      FC_W[1,14] := 0.00180894;
      FC_W[1,15] := -1.01147878;
      FC_W[1,16] := 0.31076741;
      FC_W[1,17] := -0.42154586;
      FC_W[1,18] := -0.05431300;
      FC_W[1,19] := 0.68237108;
      FC_W[1,20] := -2.56503296;
      FC_W[1,21] := 0.50673449;
      FC_W[1,22] := 0.31768897;
      FC_W[1,23] := -0.43834999;
      FC_W[1,24] := 1.20007265;
      FC_W[1,25] := 0.30830422;
      FC_W[1,26] := 0.13145778;
      FC_W[1,27] := 0.41129708;
      FC_W[1,28] := -0.09861557;
      FC_W[1,29] := -0.05401544;
      FC_W[1,30] := -0.38849521;
      FC_W[1,31] := -1.97921050;
      FC_W[2,0] := -0.79939067;
      FC_W[2,1] := 0.10302242;
      FC_W[2,2] := 0.09020624;
      FC_W[2,3] := -0.46045631;
      FC_W[2,4] := 0.32426205;
      FC_W[2,5] := 0.07683180;
      FC_W[2,6] := 0.54684573;
      FC_W[2,7] := 1.87505293;
      FC_W[2,8] := -0.48562393;
      FC_W[2,9] := 0.99263871;
      FC_W[2,10] := -0.65771282;
      FC_W[2,11] := 0.72155434;
      FC_W[2,12] := -0.66074061;
      FC_W[2,13] := 0.11306432;
      FC_W[2,14] := -0.38545227;
      FC_W[2,15] := 0.16300759;
      FC_W[2,16] := -0.02957736;
      FC_W[2,17] := -0.82533288;
      FC_W[2,18] := 0.33957723;
      FC_W[2,19] := -0.78074455;
      FC_W[2,20] := 0.55624270;
      FC_W[2,21] := -0.52731699;
      FC_W[2,22] := -1.25810063;
      FC_W[2,23] := -0.21556486;
      FC_W[2,24] := -0.03355473;
      FC_W[2,25] := 0.02170837;
      FC_W[2,26] := -0.12119742;
      FC_W[2,27] := -0.88717794;
      FC_W[2,28] := -0.91240627;
      FC_W[2,29] := 0.36170098;
      FC_W[2,30] := 0.16164558;
      FC_W[2,31] := 0.99094546;
      FC_W[3,0] := 0.19523349;
      FC_W[3,1] := 0.31197101;
      FC_W[3,2] := -0.48878455;
      FC_W[3,3] := 0.14373684;
      FC_W[3,4] := 0.24886017;
      FC_W[3,5] := -0.42134193;
      FC_W[3,6] := -0.14882350;
      FC_W[3,7] := 0.79451615;
      FC_W[3,8] := -0.46309730;
      FC_W[3,9] := 0.40033284;
      FC_W[3,10] := -0.68702614;
      FC_W[3,11] := -0.29239723;
      FC_W[3,12] := 0.98389262;
      FC_W[3,13] := 0.30846006;
      FC_W[3,14] := -0.12699004;
      FC_W[3,15] := 1.25244427;
      FC_W[3,16] := 0.17832240;
      FC_W[3,17] := -0.43285766;
      FC_W[3,18] := 0.26159754;
      FC_W[3,19] := 0.15949164;
      FC_W[3,20] := 1.06185210;
      FC_W[3,21] := 0.14212017;
      FC_W[3,22] := 0.00880439;
      FC_W[3,23] := -0.36065376;
      FC_W[3,24] := -0.39496204;
      FC_W[3,25] := -0.00392890;
      FC_W[3,26] := -0.77206844;
      FC_W[3,27] := -0.12771720;
      FC_W[3,28] := 0.72197872;
      FC_W[3,29] := 0.24183723;
      FC_W[3,30] := -0.38839531;
      FC_W[3,31] := 0.04649191;
      FC_W[4,0] := -0.42976218;
      FC_W[4,1] := 0.71019524;
      FC_W[4,2] := 0.02715457;
      FC_W[4,3] := 0.20727751;
      FC_W[4,4] := 0.12750632;
      FC_W[4,5] := 0.10362761;
      FC_W[4,6] := 0.56926334;
      FC_W[4,7] := 0.33267853;
      FC_W[4,8] := 0.22530533;
      FC_W[4,9] := -0.76057816;
      FC_W[4,10] := 0.06259055;
      FC_W[4,11] := 0.65855861;
      FC_W[4,12] := 0.43817779;
      FC_W[4,13] := -1.45052433;
      FC_W[4,14] := -0.69694483;
      FC_W[4,15] := 0.39829472;
      FC_W[4,16] := 0.00987289;
      FC_W[4,17] := 0.68149745;
      FC_W[4,18] := -0.59120047;
      FC_W[4,19] := 0.11526035;
      FC_W[4,20] := -0.45347911;
      FC_W[4,21] := 0.55277812;
      FC_W[4,22] := -0.36495659;
      FC_W[4,23] := -0.65428317;
      FC_W[4,24] := -2.59415770;
      FC_W[4,25] := 0.01274597;
      FC_W[4,26] := -0.42365780;
      FC_W[4,27] := 0.38587591;
      FC_W[4,28] := 0.33021146;
      FC_W[4,29] := 0.45073530;
      FC_W[4,30] := -0.22007711;
      FC_W[4,31] := 0.46025163;
      FC_W[5,0] := 0.08847263;
      FC_W[5,1] := 2.92971921;
      FC_W[5,2] := 0.40630540;
      FC_W[5,3] := -0.18477380;
      FC_W[5,4] := -0.35985741;
      FC_W[5,5] := 0.16343132;
      FC_W[5,6] := -1.01463449;
      FC_W[5,7] := -0.19884980;
      FC_W[5,8] := 0.19642729;
      FC_W[5,9] := 0.07467357;
      FC_W[5,10] := -0.20739354;
      FC_W[5,11] := -0.32682586;
      FC_W[5,12] := -0.24732944;
      FC_W[5,13] := -0.28553879;
      FC_W[5,14] := 0.02577983;
      FC_W[5,15] := -0.35895699;
      FC_W[5,16] := 0.13909405;
      FC_W[5,17] := -0.85842067;
      FC_W[5,18] := 0.29272711;
      FC_W[5,19] := 0.14367910;
      FC_W[5,20] := -0.33554327;
      FC_W[5,21] := -0.10857771;
      FC_W[5,22] := 0.06511363;
      FC_W[5,23] := 1.53560221;
      FC_W[5,24] := 0.36751866;
      FC_W[5,25] := 0.14096503;
      FC_W[5,26] := 0.68856186;
      FC_W[5,27] := -0.00372456;
      FC_W[5,28] := 0.07267709;
      FC_W[5,29] := 0.29737416;
      FC_W[5,30] := 0.05855417;
      FC_W[5,31] := 0.18817970;
      FC_W[6,0] := 0.22961207;
      FC_W[6,1] := 1.10309398;
      FC_W[6,2] := 1.14253712;
      FC_W[6,3] := -0.24431218;
      FC_W[6,4] := 0.24880899;
      FC_W[6,5] := 0.10031620;
      FC_W[6,6] := -1.37900984;
      FC_W[6,7] := -0.46621767;
      FC_W[6,8] := 0.23081133;
      FC_W[6,9] := -0.62265766;
      FC_W[6,10] := -0.19415495;
      FC_W[6,11] := 0.24065939;
      FC_W[6,12] := -0.37324443;
      FC_W[6,13] := 0.04941022;
      FC_W[6,14] := -0.58380717;
      FC_W[6,15] := 0.29722652;
      FC_W[6,16] := 0.45706749;
      FC_W[6,17] := 0.79749161;
      FC_W[6,18] := 0.24645862;
      FC_W[6,19] := -0.69690132;
      FC_W[6,20] := 0.25755104;
      FC_W[6,21] := -1.28122711;
      FC_W[6,22] := -0.90884095;
      FC_W[6,23] := -1.13884628;
      FC_W[6,24] := 0.61092412;
      FC_W[6,25] := 0.10356417;
      FC_W[6,26] := -0.16909865;
      FC_W[6,27] := -0.64685744;
      FC_W[6,28] := 0.09836304;
      FC_W[6,29] := 0.29990685;
      FC_W[6,30] := -0.26579708;
      FC_W[6,31] := -0.09385087;
      FC_W[7,0] := 0.11735278;
      FC_W[7,1] := 0.69732809;
      FC_W[7,2] := -0.28756016;
      FC_W[7,3] := -0.12583709;
      FC_W[7,4] := -0.44791237;
      FC_W[7,5] := 0.04257831;
      FC_W[7,6] := 0.01414247;
      FC_W[7,7] := 0.31274548;
      FC_W[7,8] := -0.42705598;
      FC_W[7,9] := 0.25311053;
      FC_W[7,10] := -0.02971629;
      FC_W[7,11] := 0.08217675;
      FC_W[7,12] := 1.13895476;
      FC_W[7,13] := 0.28638309;
      FC_W[7,14] := 0.30324531;
      FC_W[7,15] := 1.06351733;
      FC_W[7,16] := -0.09911025;
      FC_W[7,17] := -0.12825158;
      FC_W[7,18] := -0.21037468;
      FC_W[7,19] := -0.15125044;
      FC_W[7,20] := 1.04692757;
      FC_W[7,21] := -0.19273317;
      FC_W[7,22] := -0.01566108;
      FC_W[7,23] := -0.82813007;
      FC_W[7,24] := -0.17457560;
      FC_W[7,25] := -0.23310129;
      FC_W[7,26] := -0.67900503;
      FC_W[7,27] := -0.00216983;
      FC_W[7,28] := -0.33897799;
      FC_W[7,29] := 0.23453975;
      FC_W[7,30] := 0.43223280;
      FC_W[7,31] := 0.38816142;
      FC_W[8,0] := 1.24795640;
      FC_W[8,1] := 0.16966595;
      FC_W[8,2] := -0.59130764;
      FC_W[8,3] := -1.17259443;
      FC_W[8,4] := 0.58706713;
      FC_W[8,5] := -0.50881100;
      FC_W[8,6] := -0.93378001;
      FC_W[8,7] := 1.83182466;
      FC_W[8,8] := 0.69100636;
      FC_W[8,9] := -0.18218489;
      FC_W[8,10] := 0.03764156;
      FC_W[8,11] := -0.73455888;
      FC_W[8,12] := -0.53293765;
      FC_W[8,13] := 0.35738659;
      FC_W[8,14] := 0.34333083;
      FC_W[8,15] := 0.42288589;
      FC_W[8,16] := 0.47547165;
      FC_W[8,17] := 0.63862199;
      FC_W[8,18] := 0.62496924;
      FC_W[8,19] := 0.38435844;
      FC_W[8,20] := 1.82490015;
      FC_W[8,21] := 0.90129334;
      FC_W[8,22] := -0.10840212;
      FC_W[8,23] := 0.10254918;
      FC_W[8,24] := -0.91856247;
      FC_W[8,25] := 0.00505273;
      FC_W[8,26] := -0.97525537;
      FC_W[8,27] := 1.19635546;
      FC_W[8,28] := 0.29022071;
      FC_W[8,29] := 0.81490791;
      FC_W[8,30] := -0.35306564;
      FC_W[8,31] := -0.03846764;
      FC_W[9,0] := 0.53101271;
      FC_W[9,1] := 0.67765594;
      FC_W[9,2] := -0.31747413;
      FC_W[9,3] := -0.61590499;
      FC_W[9,4] := -0.35415921;
      FC_W[9,5] := 0.04045775;
      FC_W[9,6] := -0.25351635;
      FC_W[9,7] := 0.61500031;
      FC_W[9,8] := -0.00759591;
      FC_W[9,9] := 0.01995997;
      FC_W[9,10] := 0.31222284;
      FC_W[9,11] := -0.03113513;
      FC_W[9,12] := 0.55826259;
      FC_W[9,13] := 0.29481170;
      FC_W[9,14] := 0.50861734;
      FC_W[9,15] := 0.74235141;
      FC_W[9,16] := 0.04826086;
      FC_W[9,17] := 0.32700640;
      FC_W[9,18] := -0.14947560;
      FC_W[9,19] := -0.14729200;
      FC_W[9,20] := 1.31701505;
      FC_W[9,21] := 0.06887171;
      FC_W[9,22] := -0.09508032;
      FC_W[9,23] := -0.69279194;
      FC_W[9,24] := -0.32143742;
      FC_W[9,25] := -0.23362400;
      FC_W[9,26] := -0.77252012;
      FC_W[9,27] := 0.48929808;
      FC_W[9,28] := -0.59472609;
      FC_W[9,29] := 0.44059590;
      FC_W[9,30] := 0.51598865;
      FC_W[9,31] := 0.40399224;
      FC_W[10,0] := -0.05485313;
      FC_W[10,1] := 0.79143423;
      FC_W[10,2] := -0.47971761;
      FC_W[10,3] := -0.42792881;
      FC_W[10,4] := 0.76965564;
      FC_W[10,5] := 0.38477486;
      FC_W[10,6] := 0.42768925;
      FC_W[10,7] := 0.28604057;
      FC_W[10,8] := -1.25346828;
      FC_W[10,9] := 0.49736726;
      FC_W[10,10] := 0.69473928;
      FC_W[10,11] := 0.79891783;
      FC_W[10,12] := 0.62251019;
      FC_W[10,13] := 0.17432037;
      FC_W[10,14] := 1.53301835;
      FC_W[10,15] := 0.93965453;
      FC_W[10,16] := -0.46999088;
      FC_W[10,17] := 0.77361441;
      FC_W[10,18] := 0.22307561;
      FC_W[10,19] := -1.36293745;
      FC_W[10,20] := 0.20648916;
      FC_W[10,21] := 0.06673018;
      FC_W[10,22] := 0.22559744;
      FC_W[10,23] := 0.43268546;
      FC_W[10,24] := -0.21780904;
      FC_W[10,25] := -0.78115875;
      FC_W[10,26] := -0.24076101;
      FC_W[10,27] := 0.62123424;
      FC_W[10,28] := 0.29939529;
      FC_W[10,29] := 0.09014255;
      FC_W[10,30] := 0.25302246;
      FC_W[10,31] := -0.03954656;
      FC_W[11,0] := -0.24293564;
      FC_W[11,1] := -0.04531259;
      FC_W[11,2] := 0.00998670;
      FC_W[11,3] := 0.19956830;
      FC_W[11,4] := -0.20174095;
      FC_W[11,5] := -0.11596463;
      FC_W[11,6] := -0.22455990;
      FC_W[11,7] := -0.11557520;
      FC_W[11,8] := 0.41246292;
      FC_W[11,9] := 0.08150622;
      FC_W[11,10] := -1.95139670;
      FC_W[11,11] := -0.45480672;
      FC_W[11,12] := -0.08829422;
      FC_W[11,13] := 0.05833782;
      FC_W[11,14] := 0.26944444;
      FC_W[11,15] := 0.21539681;
      FC_W[11,16] := 2.23111510;
      FC_W[11,17] := 0.66294128;
      FC_W[11,18] := -0.05759437;
      FC_W[11,19] := -0.41524842;
      FC_W[11,20] := -0.13926855;
      FC_W[11,21] := 0.04841401;
      FC_W[11,22] := -0.05950727;
      FC_W[11,23] := 0.11197530;
      FC_W[11,24] := -0.04123791;
      FC_W[11,25] := -0.26082167;
      FC_W[11,26] := -0.45694438;
      FC_W[11,27] := 0.20621511;
      FC_W[11,28] := -0.53152508;
      FC_W[11,29] := 0.38166457;
      FC_W[11,30] := 0.31593123;
      FC_W[11,31] := 0.02903810;
      FC_W[12,0] := -0.11749745;
      FC_W[12,1] := -0.23415545;
      FC_W[12,2] := -0.34946913;
      FC_W[12,3] := 0.53356487;
      FC_W[12,4] := 0.18837753;
      FC_W[12,5] := -0.70393479;
      FC_W[12,6] := -0.50469047;
      FC_W[12,7] := -0.43645567;
      FC_W[12,8] := 0.66334420;
      FC_W[12,9] := -0.32834104;
      FC_W[12,10] := -1.24227428;
      FC_W[12,11] := -0.34643209;
      FC_W[12,12] := -0.28256458;
      FC_W[12,13] := -0.03548216;
      FC_W[12,14] := -0.02313955;
      FC_W[12,15] := 1.09937835;
      FC_W[12,16] := 1.40113294;
      FC_W[12,17] := 0.21808513;
      FC_W[12,18] := 0.18139383;
      FC_W[12,19] := -0.08548864;
      FC_W[12,20] := -0.56923884;
      FC_W[12,21] := 0.65053141;
      FC_W[12,22] := -0.65991580;
      FC_W[12,23] := 0.23657089;
      FC_W[12,24] := 0.02915133;
      FC_W[12,25] := -0.37136909;
      FC_W[12,26] := -0.20713671;
      FC_W[12,27] := 0.04201923;
      FC_W[12,28] := -0.21818402;
      FC_W[12,29] := 0.43879950;
      FC_W[12,30] := 0.66941983;
      FC_W[12,31] := 0.77976692;
      FC_W[13,0] := 0.05367998;
      FC_W[13,1] := 1.02593648;
      FC_W[13,2] := -1.72975278;
      FC_W[13,3] := 0.80966431;
      FC_W[13,4] := 0.03437574;
      FC_W[13,5] := -1.25336730;
      FC_W[13,6] := -0.54343611;
      FC_W[13,7] := -0.76846027;
      FC_W[13,8] := -0.07641880;
      FC_W[13,9] := -0.21239853;
      FC_W[13,10] := -1.32163453;
      FC_W[13,11] := 0.67327833;
      FC_W[13,12] := -1.27367902;
      FC_W[13,13] := -0.86751330;
      FC_W[13,14] := 0.55482459;
      FC_W[13,15] := -1.92334485;
      FC_W[13,16] := 0.08597323;
      FC_W[13,17] := -0.23974323;
      FC_W[13,18] := 0.09139446;
      FC_W[13,19] := 0.03227244;
      FC_W[13,20] := -0.22558706;
      FC_W[13,21] := -0.00554077;
      FC_W[13,22] := -0.24220449;
      FC_W[13,23] := -0.93250173;
      FC_W[13,24] := 1.33914196;
      FC_W[13,25] := -0.14073664;
      FC_W[13,26] := 1.38821757;
      FC_W[13,27] := -0.63530439;
      FC_W[13,28] := 0.86958200;
      FC_W[13,29] := -1.50805593;
      FC_W[13,30] := -0.21380891;
      FC_W[13,31] := 0.41014621;
      FC_W[14,0] := -0.63119894;
      FC_W[14,1] := -0.10577224;
      FC_W[14,2] := -0.08785659;
      FC_W[14,3] := -0.51354879;
      FC_W[14,4] := 0.30728057;
      FC_W[14,5] := -0.94762784;
      FC_W[14,6] := -0.00680102;
      FC_W[14,7] := 0.46720606;
      FC_W[14,8] := 2.24362016;
      FC_W[14,9] := -1.06858647;
      FC_W[14,10] := -1.56347978;
      FC_W[14,11] := -1.45889282;
      FC_W[14,12] := 0.46342093;
      FC_W[14,13] := 0.01371147;
      FC_W[14,14] := -0.43850195;
      FC_W[14,15] := -0.26042199;
      FC_W[14,16] := -2.62758970;
      FC_W[14,17] := -0.29780927;
      FC_W[14,18] := -1.96324050;
      FC_W[14,19] := -4.90748167;
      FC_W[14,20] := -0.20483738;
      FC_W[14,21] := -0.03886629;
      FC_W[14,22] := 1.46648896;
      FC_W[14,23] := 0.15051331;
      FC_W[14,24] := -0.04148193;
      FC_W[14,25] := -1.55939674;
      FC_W[14,26] := -0.01877716;
      FC_W[14,27] := -0.32644957;
      FC_W[14,28] := -0.03895755;
      FC_W[14,29] := -0.03125083;
      FC_W[14,30] := 0.01780568;
      FC_W[14,31] := -0.54571784;
      FC_W[15,0] := -0.89153206;
      FC_W[15,1] := 0.20046420;
      FC_W[15,2] := -0.15894163;
      FC_W[15,3] := -0.62003499;
      FC_W[15,4] := 0.67500734;
      FC_W[15,5] := -0.81095988;
      FC_W[15,6] := -0.43512601;
      FC_W[15,7] := 0.08051200;
      FC_W[15,8] := 0.22382137;
      FC_W[15,9] := 0.21324296;
      FC_W[15,10] := -1.19856393;
      FC_W[15,11] := -0.23485571;
      FC_W[15,12] := 0.08108855;
      FC_W[15,13] := -0.00869130;
      FC_W[15,14] := 0.20973921;
      FC_W[15,15] := -0.42064503;
      FC_W[15,16] := 0.83993143;
      FC_W[15,17] := 0.39107731;
      FC_W[15,18] := 0.05626461;
      FC_W[15,19] := 0.43600541;
      FC_W[15,20] := -0.40640157;
      FC_W[15,21] := -0.41479343;
      FC_W[15,22] := 1.18510294;
      FC_W[15,23] := 0.01747333;
      FC_W[15,24] := 0.27544057;
      FC_W[15,25] := 1.41735625;
      FC_W[15,26] := -1.28652883;
      FC_W[15,27] := -0.30560207;
      FC_W[15,28] := 0.28828090;
      FC_W[15,29] := 0.34294400;
      FC_W[15,30] := 1.56105816;
      FC_W[15,31] := 0.66715974;
      FC_W[16,0] := 0.18511236;
      FC_W[16,1] := 0.11142320;
      FC_W[16,2] := 0.25088802;
      FC_W[16,3] := 0.24562232;
      FC_W[16,4] := 0.23386742;
      FC_W[16,5] := 1.43394780;
      FC_W[16,6] := 1.17761219;
      FC_W[16,7] := -0.49213803;
      FC_W[16,8] := 1.12759876;
      FC_W[16,9] := 1.29781663;
      FC_W[16,10] := 0.37763405;
      FC_W[16,11] := -0.60559410;
      FC_W[16,12] := -0.58088464;
      FC_W[16,13] := -0.03103711;
      FC_W[16,14] := -0.37153244;
      FC_W[16,15] := 0.14177552;
      FC_W[16,16] := 0.08989498;
      FC_W[16,17] := -1.21121275;
      FC_W[16,18] := -1.52446818;
      FC_W[16,19] := -0.15327719;
      FC_W[16,20] := 1.36897111;
      FC_W[16,21] := -0.97303110;
      FC_W[16,22] := -1.61964941;
      FC_W[16,23] := -0.45303893;
      FC_W[16,24] := 0.07086476;
      FC_W[16,25] := -0.20691338;
      FC_W[16,26] := 0.56280392;
      FC_W[16,27] := 1.59726894;
      FC_W[16,28] := 3.60174441;
      FC_W[16,29] := -0.53792644;
      FC_W[16,30] := 2.29794812;
      FC_W[16,31] := -1.52492857;
      FC_W[17,0] := -1.34601951;
      FC_W[17,1] := -0.13013357;
      FC_W[17,2] := -0.39320931;
      FC_W[17,3] := -1.76083004;
      FC_W[17,4] := -0.25579280;
      FC_W[17,5] := -0.24240695;
      FC_W[17,6] := 0.40721077;
      FC_W[17,7] := -0.23947778;
      FC_W[17,8] := 0.50300777;
      FC_W[17,9] := -0.12915973;
      FC_W[17,10] := 3.87150478;
      FC_W[17,11] := 1.48434913;
      FC_W[17,12] := -0.27643603;
      FC_W[17,13] := 0.04503229;
      FC_W[17,14] := -0.24153562;
      FC_W[17,15] := -0.34765482;
      FC_W[17,16] := 2.79668903;
      FC_W[17,17] := -1.82834053;
      FC_W[17,18] := 0.14369456;
      FC_W[17,19] := -1.00946081;
      FC_W[17,20] := -0.00381559;
      FC_W[17,21] := -0.28470948;
      FC_W[17,22] := 1.05944335;
      FC_W[17,23] := -0.67969865;
      FC_W[17,24] := -0.14137584;
      FC_W[17,25] := -2.10863733;
      FC_W[17,26] := -1.15032828;
      FC_W[17,27] := -1.23356271;
      FC_W[17,28] := 1.35488796;
      FC_W[17,29] := 0.23205599;
      FC_W[17,30] := -0.94899446;
      FC_W[17,31] := 0.21759105;
      FC_W[18,0] := -0.86723298;
      FC_W[18,1] := 0.75922298;
      FC_W[18,2] := -0.67261380;
      FC_W[18,3] := -0.43649900;
      FC_W[18,4] := -0.02853692;
      FC_W[18,5] := 0.34614712;
      FC_W[18,6] := 0.19539559;
      FC_W[18,7] := -2.34878230;
      FC_W[18,8] := -0.42542830;
      FC_W[18,9] := 0.25120163;
      FC_W[18,10] := -1.87246346;
      FC_W[18,11] := 0.67788774;
      FC_W[18,12] := -2.58651853;
      FC_W[18,13] := 0.20881239;
      FC_W[18,14] := -0.21432896;
      FC_W[18,15] := 0.79623473;
      FC_W[18,16] := -0.35303968;
      FC_W[18,17] := -1.02341413;
      FC_W[18,18] := 0.55999649;
      FC_W[18,19] := 0.07766200;
      FC_W[18,20] := 0.00875785;
      FC_W[18,21] := 0.27602637;
      FC_W[18,22] := -0.58590114;
      FC_W[18,23] := -0.90909314;
      FC_W[18,24] := -0.31122300;
      FC_W[18,25] := -0.29507470;
      FC_W[18,26] := -3.63794160;
      FC_W[18,27] := 1.00123441;
      FC_W[18,28] := -0.59514475;
      FC_W[18,29] := 2.48554730;
      FC_W[18,30] := -0.69474798;
      FC_W[18,31] := 0.23106213;
      FC_W[19,0] := -0.11451103;
      FC_W[19,1] := -0.09549186;
      FC_W[19,2] := -0.09730008;
      FC_W[19,3] := 0.11854029;
      FC_W[19,4] := -0.33437249;
      FC_W[19,5] := -1.63624847;
      FC_W[19,6] := 0.23903780;
      FC_W[19,7] := 0.33875504;
      FC_W[19,8] := -0.75360364;
      FC_W[19,9] := -0.94568074;
      FC_W[19,10] := -0.36400679;
      FC_W[19,11] := 0.32802689;
      FC_W[19,12] := 0.33577380;
      FC_W[19,13] := -0.05023296;
      FC_W[19,14] := -0.10998800;
      FC_W[19,15] := -0.28455681;
      FC_W[19,16] := 1.20575917;
      FC_W[19,17] := -0.13861203;
      FC_W[19,18] := 1.12081277;
      FC_W[19,19] := -0.68863261;
      FC_W[19,20] := -0.53662133;
      FC_W[19,21] := -0.64450079;
      FC_W[19,22] := -0.10931280;
      FC_W[19,23] := 0.24804120;
      FC_W[19,24] := 0.19847371;
      FC_W[19,25] := -0.64389402;
      FC_W[19,26] := -0.26537114;
      FC_W[19,27] := 0.72062129;
      FC_W[19,28] := -0.21949142;
      FC_W[19,29] := 0.17651653;
      FC_W[19,30] := 0.78190112;
      FC_W[19,31] := -1.13649452;
      FC_W[20,0] := 0.83655691;
      FC_W[20,1] := 0.09223625;
      FC_W[20,2] := 0.01427277;
      FC_W[20,3] := 0.35512590;
      FC_W[20,4] := 0.29080695;
      FC_W[20,5] := -0.28151488;
      FC_W[20,6] := 2.49135256;
      FC_W[20,7] := -0.01548919;
      FC_W[20,8] := 0.31601402;
      FC_W[20,9] := -0.36315429;
      FC_W[20,10] := 0.12557349;
      FC_W[20,11] := -0.76053280;
      FC_W[20,12] := -0.00581442;
      FC_W[20,13] := 0.04770271;
      FC_W[20,14] := 0.16864912;
      FC_W[20,15] := -0.23344296;
      FC_W[20,16] := 0.58960861;
      FC_W[20,17] := 0.00711021;
      FC_W[20,18] := 0.27118811;
      FC_W[20,19] := 0.03771808;
      FC_W[20,20] := -0.36084047;
      FC_W[20,21] := 0.80696052;
      FC_W[20,22] := 0.37349138;
      FC_W[20,23] := -0.16872540;
      FC_W[20,24] := -0.27626178;
      FC_W[20,25] := 0.16081053;
      FC_W[20,26] := -0.34265164;
      FC_W[20,27] := -0.02760577;
      FC_W[20,28] := -0.31053385;
      FC_W[20,29] := -0.22049831;
      FC_W[20,30] := -0.12613228;
      FC_W[20,31] := 0.48727357;
      FC_W[21,0] := -0.29110393;
      FC_W[21,1] := 0.01953696;
      FC_W[21,2] := 0.67426211;
      FC_W[21,3] := 0.15098298;
      FC_W[21,4] := 0.25071040;
      FC_W[21,5] := 0.22902717;
      FC_W[21,6] := -1.42674541;
      FC_W[21,7] := -0.09156393;
      FC_W[21,8] := -0.76005584;
      FC_W[21,9] := -0.06921285;
      FC_W[21,10] := 0.06564474;
      FC_W[21,11] := -0.30735657;
      FC_W[21,12] := -0.29343417;
      FC_W[21,13] := 2.36240745;
      FC_W[21,14] := -0.24766001;
      FC_W[21,15] := 0.45826235;
      FC_W[21,16] := 0.58946574;
      FC_W[21,17] := -0.60599393;
      FC_W[21,18] := -0.47653148;
      FC_W[21,19] := -0.41717535;
      FC_W[21,20] := -0.14760819;
      FC_W[21,21] := 0.21080713;
      FC_W[21,22] := -0.01385766;
      FC_W[21,23] := -0.40159428;
      FC_W[21,24] := -0.53794694;
      FC_W[21,25] := 0.14114229;
      FC_W[21,26] := 0.07588908;
      FC_W[21,27] := 0.50379467;
      FC_W[21,28] := -0.29848596;
      FC_W[21,29] := -0.56126761;
      FC_W[21,30] := 0.10516994;
      FC_W[21,31] := -0.34459844;
      FC_W[22,0] := 0.50324452;
      FC_W[22,1] := -0.01163468;
      FC_W[22,2] := 0.08317020;
      FC_W[22,3] := 1.35425305;
      FC_W[22,4] := 1.03270876;
      FC_W[22,5] := 0.08969304;
      FC_W[22,6] := -0.07556182;
      FC_W[22,7] := 0.27335572;
      FC_W[22,8] := -0.06994771;
      FC_W[22,9] := -1.05795527;
      FC_W[22,10] := -0.49602944;
      FC_W[22,11] := 1.06577182;
      FC_W[22,12] := 0.24788068;
      FC_W[22,13] := -0.05016525;
      FC_W[22,14] := -0.22969624;
      FC_W[22,15] := -0.54360723;
      FC_W[22,16] := 1.10354900;
      FC_W[22,17] := -0.50223601;
      FC_W[22,18] := -1.18764758;
      FC_W[22,19] := 0.40311170;
      FC_W[22,20] := 0.27212614;
      FC_W[22,21] := -0.07391455;
      FC_W[22,22] := 0.33505601;
      FC_W[22,23] := -0.17453083;
      FC_W[22,24] := 0.07979892;
      FC_W[22,25] := -0.36740017;
      FC_W[22,26] := -0.34717765;
      FC_W[22,27] := 0.34005153;
      FC_W[22,28] := -0.45797214;
      FC_W[22,29] := -0.33705583;
      FC_W[22,30] := 0.14880560;
      FC_W[22,31] := -0.02784172;
      FC_W[23,0] := 0.89183223;
      FC_W[23,1] := 0.18917838;
      FC_W[23,2] := -0.91545367;
      FC_W[23,3] := 1.02677226;
      FC_W[23,4] := 0.67053884;
      FC_W[23,5] := 0.19384260;
      FC_W[23,6] := 0.27192867;
      FC_W[23,7] := 0.11357349;
      FC_W[23,8] := -0.85358751;
      FC_W[23,9] := 0.02984146;
      FC_W[23,10] := -0.35038522;
      FC_W[23,11] := -0.47657296;
      FC_W[23,12] := -0.20840850;
      FC_W[23,13] := -0.89233679;
      FC_W[23,14] := 0.50596559;
      FC_W[23,15] := -1.64808702;
      FC_W[23,16] := 0.83202249;
      FC_W[23,17] := -0.41169617;
      FC_W[23,18] := -0.20278446;
      FC_W[23,19] := -0.80263168;
      FC_W[23,20] := 0.08792833;
      FC_W[23,21] := 0.01297861;
      FC_W[23,22] := 0.85057580;
      FC_W[23,23] := -0.87307191;
      FC_W[23,24] := 1.66429377;
      FC_W[23,25] := 0.06264384;
      FC_W[23,26] := 2.86239386;
      FC_W[23,27] := -0.09502731;
      FC_W[23,28] := 0.38575169;
      FC_W[23,29] := 1.88736570;
      FC_W[23,30] := 0.01345321;
      FC_W[23,31] := 0.53770506;
      FC_W[24,0] := 0.21574637;
      FC_W[24,1] := 0.07279200;
      FC_W[24,2] := 0.44050846;
      FC_W[24,3] := 1.07333148;
      FC_W[24,4] := 1.29573095;
      FC_W[24,5] := -0.01340208;
      FC_W[24,6] := -0.01077834;
      FC_W[24,7] := 0.43822077;
      FC_W[24,8] := -0.13799220;
      FC_W[24,9] := -1.20653403;
      FC_W[24,10] := -0.66901463;
      FC_W[24,11] := 0.65269983;
      FC_W[24,12] := 0.37482554;
      FC_W[24,13] := 0.01565100;
      FC_W[24,14] := 0.12979744;
      FC_W[24,15] := -0.87315303;
      FC_W[24,16] := 0.69985312;
      FC_W[24,17] := -0.31910187;
      FC_W[24,18] := -1.57823551;
      FC_W[24,19] := 1.63719082;
      FC_W[24,20] := 0.53801286;
      FC_W[24,21] := -0.89269280;
      FC_W[24,22] := 0.43086779;
      FC_W[24,23] := -0.36367694;
      FC_W[24,24] := 0.13592418;
      FC_W[24,25] := -1.06909513;
      FC_W[24,26] := -0.36003765;
      FC_W[24,27] := 0.18487933;
      FC_W[24,28] := -0.71037912;
      FC_W[24,29] := -0.13214959;
      FC_W[24,30] := 0.38270515;
      FC_W[24,31] := -0.22937216;
      FC_W[25,0] := 0.22048582;
      FC_W[25,1] := 0.07118796;
      FC_W[25,2] := 0.43118235;
      FC_W[25,3] := 1.09670317;
      FC_W[25,4] := 1.30268395;
      FC_W[25,5] := -0.02062076;
      FC_W[25,6] := -0.00384964;
      FC_W[25,7] := 0.42397165;
      FC_W[25,8] := -0.13090287;
      FC_W[25,9] := -1.19230533;
      FC_W[25,10] := -0.64925510;
      FC_W[25,11] := 0.66327566;
      FC_W[25,12] := 0.36542091;
      FC_W[25,13] := 0.01464875;
      FC_W[25,14] := 0.11140072;
      FC_W[25,15] := -0.85105401;
      FC_W[25,16] := 0.71580303;
      FC_W[25,17] := -0.31853670;
      FC_W[25,18] := -1.57619953;
      FC_W[25,19] := 1.59803832;
      FC_W[25,20] := 0.52842081;
      FC_W[25,21] := -0.88470274;
      FC_W[25,22] := 0.43769893;
      FC_W[25,23] := -0.35991374;
      FC_W[25,24] := 0.13580397;
      FC_W[25,25] := -1.04141033;
      FC_W[25,26] := -0.34737530;
      FC_W[25,27] := 0.18887003;
      FC_W[25,28] := -0.71740890;
      FC_W[25,29] := -0.13793097;
      FC_W[25,30] := 0.37530687;
      FC_W[25,31] := -0.23953751;
      FC_W[26,0] := 1.56152236;
      FC_W[26,1] := 0.10283720;
      FC_W[26,2] := -1.14192486;
      FC_W[26,3] := 0.12904538;
      FC_W[26,4] := 0.07129417;
      FC_W[26,5] := -0.00974355;
      FC_W[26,6] := 0.26723784;
      FC_W[26,7] := 0.26951763;
      FC_W[26,8] := -0.80771482;
      FC_W[26,9] := -0.63183504;
      FC_W[26,10] := -0.73038095;
      FC_W[26,11] := 0.70714259;
      FC_W[26,12] := 0.49866056;
      FC_W[26,13] := -1.70901299;
      FC_W[26,14] := -0.73239201;
      FC_W[26,15] := -1.52383792;
      FC_W[26,16] := 1.03083646;
      FC_W[26,17] := 0.14269158;
      FC_W[26,18] := -0.67796141;
      FC_W[26,19] := -0.46712342;
      FC_W[26,20] := -0.29322225;
      FC_W[26,21] := 0.83879727;
      FC_W[26,22] := -0.64477837;
      FC_W[26,23] := 0.34093615;
      FC_W[26,24] := 0.58871043;
      FC_W[26,25] := -0.27591738;
      FC_W[26,26] := -0.80217528;
      FC_W[26,27] := -0.24964441;
      FC_W[26,28] := 0.87935400;
      FC_W[26,29] := -0.08472463;
      FC_W[26,30] := -0.02381817;
      FC_W[26,31] := 1.22797525;
      FC_W[27,0] := 0.38102069;
      FC_W[27,1] := 0.09269264;
      FC_W[27,2] := 0.59470004;
      FC_W[27,3] := 0.28748643;
      FC_W[27,4] := -0.09679463;
      FC_W[27,5] := -0.41851318;
      FC_W[27,6] := -1.15975082;
      FC_W[27,7] := 0.02223462;
      FC_W[27,8] := -0.34720707;
      FC_W[27,9] := 0.72622478;
      FC_W[27,10] := 0.11481044;
      FC_W[27,11] := 0.37256941;
      FC_W[27,12] := -0.20693421;
      FC_W[27,13] := 2.54740143;
      FC_W[27,14] := -0.02115205;
      FC_W[27,15] := 0.28944260;
      FC_W[27,16] := -0.51868707;
      FC_W[27,17] := -0.03483006;
      FC_W[27,18] := -0.59467632;
      FC_W[27,19] := 0.17160304;
      FC_W[27,20] := -0.60751998;
      FC_W[27,21] := -0.62638927;
      FC_W[27,22] := 0.10618542;
      FC_W[27,23] := -0.31771034;
      FC_W[27,24] := -0.97128564;
      FC_W[27,25] := -0.43134749;
      FC_W[27,26] := 0.02182774;
      FC_W[27,27] := -0.32529354;
      FC_W[27,28] := 0.34785143;
      FC_W[27,29] := -0.04944998;
      FC_W[27,30] := 0.33690751;
      FC_W[27,31] := 0.17198400;
      FC_W[28,0] := 0.77232850;
      FC_W[28,1] := 0.02787268;
      FC_W[28,2] := 0.41619617;
      FC_W[28,3] := 0.23172490;
      FC_W[28,4] := -0.09291978;
      FC_W[28,5] := -0.21665370;
      FC_W[28,6] := -0.98798215;
      FC_W[28,7] := -0.12977834;
      FC_W[28,8] := -0.46919557;
      FC_W[28,9] := 0.74807566;
      FC_W[28,10] := -0.13898452;
      FC_W[28,11] := -0.46674505;
      FC_W[28,12] := -0.17911388;
      FC_W[28,13] := -1.79411507;
      FC_W[28,14] := 0.06221046;
      FC_W[28,15] := 0.05005321;
      FC_W[28,16] := 0.66611379;
      FC_W[28,17] := -0.69680721;
      FC_W[28,18] := 0.19765745;
      FC_W[28,19] := -0.42630407;
      FC_W[28,20] := -0.27623644;
      FC_W[28,21] := -0.38921455;
      FC_W[28,22] := 0.35367966;
      FC_W[28,23] := -0.44775704;
      FC_W[28,24] := -1.63023448;
      FC_W[28,25] := -0.28671730;
      FC_W[28,26] := 0.01121899;
      FC_W[28,27] := 0.26976588;
      FC_W[28,28] := -0.29760954;
      FC_W[28,29] := -0.63540250;
      FC_W[28,30] := 0.43073460;
      FC_W[28,31] := 0.22689007;
      FC_W[29,0] := -0.40210408;
      FC_W[29,1] := 0.69945884;
      FC_W[29,2] := -0.76612192;
      FC_W[29,3] := 0.48992610;
      FC_W[29,4] := 2.01849413;
      FC_W[29,5] := -0.82425791;
      FC_W[29,6] := 1.45209885;
      FC_W[29,7] := -1.13971364;
      FC_W[29,8] := -0.31848440;
      FC_W[29,9] := 2.11410785;
      FC_W[29,10] := 1.93272853;
      FC_W[29,11] := -0.68537265;
      FC_W[29,12] := -1.44989634;
      FC_W[29,13] := -0.19573005;
      FC_W[29,14] := -2.68635106;
      FC_W[29,15] := 0.50114202;
      FC_W[29,16] := -0.05285606;
      FC_W[29,17] := 3.36546516;
      FC_W[29,18] := -0.43367249;
      FC_W[29,19] := 0.21831593;
      FC_W[29,20] := 0.49202019;
      FC_W[29,21] := -1.24413443;
      FC_W[29,22] := 1.24901104;
      FC_W[29,23] := 0.13342574;
      FC_W[29,24] := 0.18592642;
      FC_W[29,25] := -0.82732177;
      FC_W[29,26] := -0.10154523;
      FC_W[29,27] := 0.68388170;
      FC_W[29,28] := -1.91055167;
      FC_W[29,29] := -1.10603726;
      FC_W[29,30] := 0.22993748;
      FC_W[29,31] := -2.25390053;
      FC_W[30,0] := 0.50542051;
      FC_W[30,1] := -0.01288069;
      FC_W[30,2] := 0.07892181;
      FC_W[30,3] := 1.35607970;
      FC_W[30,4] := 1.02726829;
      FC_W[30,5] := 0.09714934;
      FC_W[30,6] := -0.07362376;
      FC_W[30,7] := 0.27333879;
      FC_W[30,8] := -0.07077026;
      FC_W[30,9] := -1.05870450;
      FC_W[30,10] := -0.49826735;
      FC_W[30,11] := 1.07048607;
      FC_W[30,12] := 0.24682963;
      FC_W[30,13] := -0.05297443;
      FC_W[30,14] := -0.23532499;
      FC_W[30,15] := -0.54376680;
      FC_W[30,16] := 1.10788131;
      FC_W[30,17] := -0.50225794;
      FC_W[30,18] := -1.18030238;
      FC_W[30,19] := 0.39142749;
      FC_W[30,20] := 0.27120695;
      FC_W[30,21] := -0.06207144;
      FC_W[30,22] := 0.33196387;
      FC_W[30,23] := -0.17185551;
      FC_W[30,24] := 0.07908980;
      FC_W[30,25] := -0.36303857;
      FC_W[30,26] := -0.35007730;
      FC_W[30,27] := 0.34561849;
      FC_W[30,28] := -0.45720354;
      FC_W[30,29] := -0.34233299;
      FC_W[30,30] := 0.14847992;
      FC_W[30,31] := -0.02407410;
      FC_W[31,0] := 0.70713001;
      FC_W[31,1] := -0.00918456;
      FC_W[31,2] := 0.11002598;
      FC_W[31,3] := 2.00804901;
      FC_W[31,4] := 0.88700664;
      FC_W[31,5] := 0.47887260;
      FC_W[31,6] := -0.14625056;
      FC_W[31,7] := 0.47002777;
      FC_W[31,8] := 0.34443581;
      FC_W[31,9] := -0.70228255;
      FC_W[31,10] := -0.85665584;
      FC_W[31,11] := 2.20079017;
      FC_W[31,12] := 0.36255807;
      FC_W[31,13] := -0.06039402;
      FC_W[31,14] := -0.22185645;
      FC_W[31,15] := -0.70947796;
      FC_W[31,16] := 0.43582395;
      FC_W[31,17] := -0.48801118;
      FC_W[31,18] := -0.39800802;
      FC_W[31,19] := 0.48426980;
      FC_W[31,20] := 0.24603498;
      FC_W[31,21] := 0.19021983;
      FC_W[31,22] := 0.91978002;
      FC_W[31,23] := -0.20594357;
      FC_W[31,24] := 0.06884714;
      FC_W[31,25] := -1.04134059;
      FC_W[31,26] := -0.62354541;
      FC_W[31,27] := 0.30330026;
      FC_W[31,28] := -0.12263997;
      FC_W[31,29] := -0.36841112;
      FC_W[31,30] := 0.44422802;
      FC_W[31,31] := 0.36350179;
      FC_W[32,0] := 0.85074222;
      FC_W[32,1] := -0.07046198;
      FC_W[32,2] := -0.00526896;
      FC_W[32,3] := 1.48461521;
      FC_W[32,4] := 0.79624808;
      FC_W[32,5] := -0.32169014;
      FC_W[32,6] := -0.02443201;
      FC_W[32,7] := 0.08702906;
      FC_W[32,8] := 0.19203611;
      FC_W[32,9] := -0.77823097;
      FC_W[32,10] := -0.18044655;
      FC_W[32,11] := 1.29543126;
      FC_W[32,12] := 0.04275373;
      FC_W[32,13] := 0.05409016;
      FC_W[32,14] := -0.23328111;
      FC_W[32,15] := -0.17099567;
      FC_W[32,16] := 1.38528931;
      FC_W[32,17] := -0.58370709;
      FC_W[32,18] := -1.28326952;
      FC_W[32,19] := -0.41117722;
      FC_W[32,20] := -0.00477389;
      FC_W[32,21] := -0.14191154;
      FC_W[32,22] := 0.11423180;
      FC_W[32,23] := -0.05158845;
      FC_W[32,24] := -0.08476931;
      FC_W[32,25] := 0.31649798;
      FC_W[32,26] := -0.12338689;
      FC_W[32,27] := 0.19256236;
      FC_W[32,28] := -0.36851650;
      FC_W[32,29] := -0.19011347;
      FC_W[32,30] := -0.14693265;
      FC_W[32,31] := -0.21090116;
      FC_W[33,0] := 1.17051291;
      FC_W[33,1] := -0.18128292;
      FC_W[33,2] := -0.24709880;
      FC_W[33,3] := 1.54797363;
      FC_W[33,4] := 0.27815264;
      FC_W[33,5] := -0.25975022;
      FC_W[33,6] := -0.18560846;
      FC_W[33,7] := -0.00064327;
      FC_W[33,8] := 0.31427521;
      FC_W[33,9] := -0.66741139;
      FC_W[33,10] := -0.11064007;
      FC_W[33,11] := 1.71599257;
      FC_W[33,12] := -0.01325114;
      FC_W[33,13] := 0.05017950;
      FC_W[33,14] := -0.33987817;
      FC_W[33,15] := 0.11878651;
      FC_W[33,16] := 1.68803883;
      FC_W[33,17] := -0.89897865;
      FC_W[33,18] := -0.86278552;
      FC_W[33,19] := -1.63729823;
      FC_W[33,20] := -0.31710440;
      FC_W[33,21] := 0.60572541;
      FC_W[33,22] := -0.15609778;
      FC_W[33,23] := 0.14094375;
      FC_W[33,24] := -0.22354113;
      FC_W[33,25] := 1.02642429;
      FC_W[33,26] := -0.13626578;
      FC_W[33,27] := 0.24193136;
      FC_W[33,28] := 0.02687795;
      FC_W[33,29] := -0.25783661;
      FC_W[33,30] := -0.42547590;
      FC_W[33,31] := 0.06487284;
      FC_W[34,0] := 0.93701762;
      FC_W[34,1] := -0.13635513;
      FC_W[34,2] := -0.14065792;
      FC_W[34,3] := 1.31602311;
      FC_W[34,4] := 0.31817526;
      FC_W[34,5] := -0.04061212;
      FC_W[34,6] := -0.24273089;
      FC_W[34,7] := 0.12358569;
      FC_W[34,8] := 0.26035085;
      FC_W[34,9] := -0.93310243;
      FC_W[34,10] := -0.31741625;
      FC_W[34,11] := 1.51594436;
      FC_W[34,12] := 0.08120698;
      FC_W[34,13] := 0.01410864;
      FC_W[34,14] := -0.17541805;
      FC_W[34,15] := -0.06809679;
      FC_W[34,16] := 1.51319253;
      FC_W[34,17] := -0.88881022;
      FC_W[34,18] := -0.84934044;
      FC_W[34,19] := -1.14595699;
      FC_W[34,20] := -0.14682929;
      FC_W[34,21] := 0.57783365;
      FC_W[34,22] := -0.15478867;
      FC_W[34,23] := 0.03422264;
      FC_W[34,24] := -0.16054711;
      FC_W[34,25] := 0.72221678;
      FC_W[34,26] := -0.22578676;
      FC_W[34,27] := 0.23727337;
      FC_W[34,28] := -0.02117160;
      FC_W[34,29] := -0.20905079;
      FC_W[34,30] := -0.29970139;
      FC_W[34,31] := 0.20462438;
      FC_W[35,0] := 0.74387974;
      FC_W[35,1] := 0.00046961;
      FC_W[35,2] := 0.12905753;
      FC_W[35,3] := 1.42334437;
      FC_W[35,4] := 1.01942086;
      FC_W[35,5] := -0.51153046;
      FC_W[35,6] := 0.09392732;
      FC_W[35,7] := 0.08796729;
      FC_W[35,8] := 0.19130485;
      FC_W[35,9] := -0.76946145;
      FC_W[35,10] := -0.12217331;
      FC_W[35,11] := 1.03380001;
      FC_W[35,12] := 0.00288362;
      FC_W[35,13] := 0.09569277;
      FC_W[35,14] := -0.11386733;
      FC_W[35,15] := -0.25902045;
      FC_W[35,16] := 1.27864158;
      FC_W[35,17] := -0.42641610;
      FC_W[35,18] := -1.57564640;
      FC_W[35,19] := 0.09335784;
      FC_W[35,20] := 0.10024387;
      FC_W[35,21] := -0.62594521;
      FC_W[35,22] := 0.19663191;
      FC_W[35,23] := -0.16496119;
      FC_W[35,24] := -0.03103490;
      FC_W[35,25] := 0.10913338;
      FC_W[35,26] := 0.03627454;
      FC_W[35,27] := 0.10267387;
      FC_W[35,28] := -0.56860989;
      FC_W[35,29] := -0.03318772;
      FC_W[35,30] := -0.08832761;
      FC_W[35,31] := -0.44099909;
      FC_W[36,0] := 0.52166957;
      FC_W[36,1] := -0.12047767;
      FC_W[36,2] := -0.65333307;
      FC_W[36,3] := 1.27468884;
      FC_W[36,4] := 0.85022986;
      FC_W[36,5] := 1.30502415;
      FC_W[36,6] := 0.51394087;
      FC_W[36,7] := -0.21489781;
      FC_W[36,8] := 0.47256544;
      FC_W[36,9] := -2.08075500;
      FC_W[36,10] := -0.15392257;
      FC_W[36,11] := -0.91717398;
      FC_W[36,12] := -0.23858869;
      FC_W[36,13] := 1.36014390;
      FC_W[36,14] := 0.04703877;
      FC_W[36,15] := 0.53182036;
      FC_W[36,16] := 0.82169122;
      FC_W[36,17] := 0.12479233;
      FC_W[36,18] := -0.55995673;
      FC_W[36,19] := 1.01603258;
      FC_W[36,20] := 0.16605985;
      FC_W[36,21] := -4.44515848;
      FC_W[36,22] := 0.33325189;
      FC_W[36,23] := 0.35819244;
      FC_W[36,24] := -1.46462762;
      FC_W[36,25] := -0.33244470;
      FC_W[36,26] := -0.22851460;
      FC_W[36,27] := -0.70994413;
      FC_W[36,28] := -1.00351298;
      FC_W[36,29] := -0.68896842;
      FC_W[36,30] := 0.19659905;
      FC_W[36,31] := 0.11465314;
      FC_W[37,0] := 0.72986430;
      FC_W[37,1] := 0.01660483;
      FC_W[37,2] := 0.15380096;
      FC_W[37,3] := 1.42001820;
      FC_W[37,4] := 1.08455575;
      FC_W[37,5] := -0.56139719;
      FC_W[37,6] := 0.11629014;
      FC_W[37,7] := 0.08233827;
      FC_W[37,8] := 0.19204774;
      FC_W[37,9] := -0.75335324;
      FC_W[37,10] := -0.10558938;
      FC_W[37,11] := 0.97539324;
      FC_W[37,12] := -0.01387812;
      FC_W[37,13] := 0.11496376;
      FC_W[37,14] := -0.09327843;
      FC_W[37,15] := -0.28244978;
      FC_W[37,16] := 1.24588180;
      FC_W[37,17] := -0.37139711;
      FC_W[37,18] := -1.65386844;
      FC_W[37,19] := 0.22961944;
      FC_W[37,20] := 0.12245397;
      FC_W[37,21] := -0.77627939;
      FC_W[37,22] := 0.22540502;
      FC_W[37,23] := -0.18894139;
      FC_W[37,24] := -0.01488678;
      FC_W[37,25] := 0.04418439;
      FC_W[37,26] := 0.06954633;
      FC_W[37,27] := 0.06961229;
      FC_W[37,28] := -0.62086546;
      FC_W[37,29] := -0.00426411;
      FC_W[37,30] := -0.06620175;
      FC_W[37,31] := -0.50101370;
      FC_W[38,0] := 1.00738335;
      FC_W[38,1] := 0.09097587;
      FC_W[38,2] := -0.22697389;
      FC_W[38,3] := 0.43213934;
      FC_W[38,4] := 0.23431744;
      FC_W[38,5] := 0.55504799;
      FC_W[38,6] := -0.46511737;
      FC_W[38,7] := -0.30007234;
      FC_W[38,8] := -0.89533710;
      FC_W[38,9] := -0.89366823;
      FC_W[38,10] := 0.45313212;
      FC_W[38,11] := 0.04846459;
      FC_W[38,12] := -0.36337411;
      FC_W[38,13] := -0.02901641;
      FC_W[38,14] := 0.02675290;
      FC_W[38,15] := 0.21207911;
      FC_W[38,16] := -1.05750823;
      FC_W[38,17] := 0.03571362;
      FC_W[38,18] := -0.54906017;
      FC_W[38,19] := -0.06487506;
      FC_W[38,20] := 1.46296978;
      FC_W[38,21] := 1.68687689;
      FC_W[38,22] := -0.79362643;
      FC_W[38,23] := 0.01360563;
      FC_W[38,24] := -0.90076172;
      FC_W[38,25] := -0.03557481;
      FC_W[38,26] := 0.01827911;
      FC_W[38,27] := -4.41204262;
      FC_W[38,28] := 1.03043067;
      FC_W[38,29] := 0.07150628;
      FC_W[38,30] := 0.89232284;
      FC_W[38,31] := -2.00459933;
      FC_W[39,0] := -1.00683630;
      FC_W[39,1] := 0.35158142;
      FC_W[39,2] := -0.14014471;
      FC_W[39,3] := 3.00387716;
      FC_W[39,4] := 0.24598759;
      FC_W[39,5] := -0.02767153;
      FC_W[39,6] := -1.18190074;
      FC_W[39,7] := 0.73443639;
      FC_W[39,8] := 1.13997531;
      FC_W[39,9] := -0.14120299;
      FC_W[39,10] := 1.32576215;
      FC_W[39,11] := -1.01461887;
      FC_W[39,12] := 0.55732387;
      FC_W[39,13] := 0.06342927;
      FC_W[39,14] := 0.90479892;
      FC_W[39,15] := -1.52994144;
      FC_W[39,16] := -0.29925072;
      FC_W[39,17] := 1.18414056;
      FC_W[39,18] := -0.38163671;
      FC_W[39,19] := -1.38458204;
      FC_W[39,20] := 0.27376747;
      FC_W[39,21] := 0.20587626;
      FC_W[39,22] := -0.30574843;
      FC_W[39,23] := -0.27512020;
      FC_W[39,24] := -0.03444282;
      FC_W[39,25] := 0.02989091;
      FC_W[39,26] := -1.41995561;
      FC_W[39,27] := -0.64386964;
      FC_W[39,28] := 1.14525557;
      FC_W[39,29] := 0.62678617;
      FC_W[39,30] := -0.04682657;
      FC_W[39,31] := 0.28188556;
      FC_B[0] := 0.27300268;
      FC_B[1] := -0.03010342;
      FC_B[2] := -0.01271929;
      FC_B[3] := 0.43827111;
      FC_B[4] := 0.13327518;
      FC_B[5] := 0.57994288;
      FC_B[6] := 0.21499516;
      FC_B[7] := -0.06454320;
      FC_B[8] := -0.32960591;
      FC_B[9] := -0.43125266;
      FC_B[10] := -0.37227541;
      FC_B[11] := 0.73980105;
      FC_B[12] := -0.20920722;
      FC_B[13] := -0.39066130;
      FC_B[14] := -0.07623728;
      FC_B[15] := -0.73917663;
      FC_B[16] := 0.42881081;
      FC_B[17] := -0.65394527;
      FC_B[18] := 0.39339224;
      FC_B[19] := -0.48604643;
      FC_B[20] := -0.11493951;
      FC_B[21] := 0.28442013;
      FC_B[22] := -1.20434070;
      FC_B[23] := -0.69569170;
      FC_B[24] := -1.20312428;
      FC_B[25] := -1.20610702;
      FC_B[26] := -1.35554242;
      FC_B[27] := 0.75533146;
      FC_B[28] := -0.01746950;
      FC_B[29] := 0.87777281;
      FC_B[30] := -1.20342910;
      FC_B[31] := -0.59860963;
      FC_B[32] := -1.29991877;
      FC_B[33] := -1.25148046;
      FC_B[34] := -1.24426150;
      FC_B[35] := -1.35175025;
      FC_B[36] := 0.02938923;
      FC_B[37] := -1.35940027;
      FC_B[38] := 1.13188744;
      FC_B[39] := 1.56624103;

END_DATA_BLOCK
